(* IEC 61131-3 sources: mapprobotics-sample-tracking/FileDevices/GCode, 6 files *)

(* ---- ProdDetails.typ ---- *)
TYPE
	ProductDetailsType : 	STRUCT  (*Additional data added as attributes to every tracking object*)
		This : UDINT; (*Adress to the memory - debugging*)
		GripperClosed : BOOL; (*Gripper is close, product in manipulation*)
		TrackingFrameID : UDINT; (*tracking frame id*)
		PickPosDelta : McPosType;
		PickPos : McPosType; (*position where gripper has been closed*)
		IncrementPos : McPosType; (*change in position on frame*)
		Pos : McPosType; (*Actual Position of object*)
		ObjectType : USINT; (*Classification of the object (red / blue)*)
		InTracking : BOOL; (*Object is now active in Tracking*)
		Robot : DevicesListEnum; (*type of robot manipulated the object*)
	END_STRUCT;
	DevicesListEnum :
		( (*device definition of manipulating robots and axis*)
		DEV_Conveyor := 0, (*object id for conveyor*)
		DEV_Robot := 1, (*id for robot 1*)
		DEV_Removed := 2 (*marked as removed and do not show in scene*)
		);
END_TYPE

(* ---- Multipick.st ---- *)
#include 'ProdDetails.typ'

////////////////////////////////////////////////////////////////////////////////////
// INPUT Variables - configured as Program Elements of the interpreter
	// NextTrackingObjectIn : UDINT;							 Pointer to next object (GCS)

// OUTPUT Variables - configured as Program Elements of the interpreter
	// MaxPickPosIn : LREAL;								 	Maximum Position where robot is able to grab something (BCS)
	// MinPickPosIn : LREAL;								 	Minimum Position where objects are given to the robot (BCS)

VAR CONSTANT
	UpperZLevel : LREAL := 100.0;	// Gripper up position
	LowerZLevel : LREAL := 0.0;		// Gripper down position
	YProductPos : LREAL := 200;		// position in y coordinate where the product should be placed
END_VAR

VAR
	ActObj 	: REFERENCE TO ProductDetailsType;
	NextObj : REFERENCE TO ProductDetailsType;
	ParkPos				: McPointType := (Pos:=(X:=	  0, Y:= 0, 			Z:= UpperZLevel));
	SynchPosUp1			: McPointType := (Pos:=(X:=   -100, Y:= 0, 			Z:= UpperZLevel));
	SynchPosUp2			: McPointType := (Pos:=(X:=   100, Y:= 0, 			Z:= UpperZLevel));
	SynchPosDown1		: McPointType := (Pos:=(X:=   -100, Y:= 0, 			Z:= LowerZLevel));
	SynchPosDown2		: McPointType := (Pos:=(X:=   100, Y:= 0, 			Z:= LowerZLevel));
	StaticMoveDown		: McPointType := (Pos:=(X:=	  0, Y:= 0, 			Z:= 0));
	MoveToPark : BOOL 	:= FALSE;
END_VAR

PROGRAM _MAIN

	// Position init, reset frame in case of restart
	SetPCS(MachineFrame);
	MoveLR(ParkPos);

	// Set the manipulation area of the Robot
	MaxPickPosIn := 1400;
	MinPickPosIn := 200;

	REPEAT
		IF NextTrackingObjectIn <> 0 THEN
			MoveToPark := FALSE;

			ActObj ACCESS NextTrackingObjectIn;								// select the product
			TrackObjectR(ActObj.TrackingFrameID, SynchPosUp2, 50, 50);		// track on product
			MoveLR(SynchPosDown2);											// move to the take position
			SetM(34);														// Scene - remove product from belt, Close the gripper here
			WaitTime(0.04);													// Wait cause delay of gripper
			WaitALAP();
			MoveLR(SynchPosUp2);											// move up to change position

			NextObj ACCESS NextTrackingObjectIn;
			IF ADR(NextObj) <> 0 AND ADR(NextObj) <> ADR(ActObj) THEN
				TrackObjectR(NextObj.TrackingFrameID, SynchPosUp1, 50, 50);	// track on product
				MoveLR(SynchPosDown1);										// move to the take position
				SetM(33);													// Scene - remove product from belt, Close the gripper here
				WaitTime(0.04);												// Wait cause delay of gripper
				MoveLR(SynchPosUp1);										// move up to change position
			END_IF

			TrackStopR(FixedPlace, ParkPos, 50, 50);						// Move to the fixed place Position
			MoveLR(StaticMoveDown);											// move to the take position
			SetM(16);														// open the gripper here
			SetM(17);														// open the gripper here
			WaitTime(0.04);													// Wait cause delay of gripper
			MoveLR(ParkPos);												// move to the take position
			WaitALAP();

			IF NextTrackingObjectIn = 0 THEN								// Need to stop, no objects left
				MoveToPark := TRUE;											// force park position
			END_IF

		ELSE
			MoveToPark := TRUE;												// force park position, there is nothing to take
		END_IF

		IF MoveToPark THEN
			MoveLR(ParkPos);												// move to static park position
			WaitEndMove();													// sync interpreter and program
			WaitIp();														// hold interpreter until a new frame is available
		END_IF

	UNTIL FALSE END_REPEAT;

END_PROGRAM

(* ---- PickNPlace.st ---- *)
#include 'ProdDetails.typ'

////////////////////////////////////////////////////////////////////////////////////
// INPUT Variables - configured as Program Elements of the interpreter
	// NextTrackingObjectIn : UDINT;							 Pointer to next object (GCS)
	// NextTrackingObjectOut : UDINT;							 Pointer to next object (GCS)

// OUTPUT Variables - configured as Program Elements of the interpreter
	// MaxPickPosIn : LREAL;								 	Maximum Position where robot is able to grab something (BCS)
	// MinPickPosIn : LREAL;								 	Minimum Position where objects are given to the robot (BCS)
	// MaxPickPosOut : LREAL;								 	Maximum Position where robot is able to place something (BCS)
	// MinPickPosOut : LREAL;								 	Minimum Position where objects are placed by the robot (BCS)

VAR CONSTANT
	UpperZLevel : LREAL := 100.0;	// Gripper up position
	LowerZLevel : LREAL := 0.0;		// Gripper down position
	YProductPos : LREAL := 200;		// position in y coordinate where the product should be placed
END_VAR

VAR
	ActObj : REFERENCE TO ProductDetailsType;
	ParkPos				: McPointType := (Pos:=(X:=-100, Y:=100, 			Z:= UpperZLevel));
	SynchPosUp			: McPointType := (Pos:=(X:=   0, Y:= 0, 			Z:= UpperZLevel));
	SynchPosDown		: McPointType := (Pos:=(X:=   0, Y:= 0, 			Z:= LowerZLevel));
	MoveToPark : BOOL := FALSE;
END_VAR

PROGRAM _MAIN

	// Position init, reset frame in case of restart
	SetPCS(MachineFrame);
	MoveLR(ParkPos);

	// Set the manipulation area of the Robot
	MaxPickPosIn := 1400;
	MinPickPosIn := 400;
	MaxPickPosOut := 1700;
	MinPickPosOut := 700;

	REPEAT
		IF NextTrackingObjectIn <> 0 THEN
			MoveToPark := FALSE;

			ActObj ACCESS NextTrackingObjectIn;							// select the product
			TrackObjectR(ActObj.TrackingFrameID, SynchPosUp, 50, 50);	// track on product
			MoveLR(SynchPosDown);										// move to the take position
			WaitALAP();													// hold interpreter
			SetM(32);													// Scene - remove product from belt, close gripper
			WaitTime(0.04);												// Wait cause delay of gripper

			MoveLR(SynchPosUp);											// move up to change frame
			WaitUntil(NextTrackingObjectOut <> 0);						// hold interpeter until place frame has been selected
			ActObj ACCESS NextTrackingObjectOut;						// change memory reference
			TrackObjectR(ActObj.TrackingFrameID, SynchPosUp, 50, 50);	// move to place position
			MoveLR(SynchPosDown);										// move down on place position
			WaitALAP();													// hold interpreter
			SetM(16);													// Scene - place product on belt, open gripper
			WaitTime(0.04);												// Wait cause delay of gripper

			MoveLR(SynchPosUp);											// move up to change frame
			IF NextTrackingObjectIn = 0 THEN							// Need to stop, no objects left
				TrackStopR(MachineFrame, ParkPos, 50, 50);				// Move to a static frame
				MoveToPark := TRUE;										// force park position
			END_IF

		ELSE
			MoveToPark := TRUE;											// force park position, there is nothing to take
		END_IF

		IF MoveToPark THEN
			MoveLR(ParkPos);											// move to static park position
			WaitEndMove();												// sync interpreter and program
			WaitIp();													// hold interpreter until a new frame is available
		END_IF

	UNTIL FALSE END_REPEAT;

END_PROGRAM

(* ---- PlaceWithConditionalStop.st ---- *)
#include 'ProdDetails.typ'

////////////////////////////////////////////////////////////////////////////////////
// INPUT Variables - configured as Program Elements of the interpreter
	// NextTrackingObjectIn : UDINT;							 Pointer to next object (GCS)

// OUTPUT Variables - configured as Program Elements of the interpreter
	// MaxPickPosIn : LREAL;								 	Maximum Position where robot is able to grab something (BCS)
	// MinPickPosIn : LREAL;								 	Minimum Position where objects are given to the robot (BCS)

VAR CONSTANT
	UpperZLevel : LREAL := 100.0;	// Gripper up position
	LowerZLevel : LREAL := 0.0;		// Gripper down position
	YProductPos : LREAL := 200;		// position in y coordinate where the product should be placed
END_VAR

VAR
	ActObj : REFERENCE TO ProductDetailsType;
	ParkPos				: McPointType := (Pos:=(X:=	  0, Y:= 0, 			Z:= UpperZLevel));
	SynchPosUp			: McPointType := (Pos:=(X:=   0, Y:= 0, 			Z:= UpperZLevel));
	SynchPosDown		: McPointType := (Pos:=(X:=   0, Y:= 0, 			Z:= LowerZLevel));
	StaticMoveDown		: McPointType := (Pos:=(X:=   0, Y:= 0, 			Z:= -100));
	StaticMoveUp		: McPointType := (Pos:=(X:=   0, Y:= 0, 			Z:= 100));
	MoveToPark : BOOL 	:= FALSE;
END_VAR

PROGRAM _MAIN

	// Position init, reset frame in case of restart
	SetPCS(MachineFrame);
	MoveLR(ParkPos);

	// Set the manipulation area of the Robot
	MaxPickPosIn := 1400;
	MinPickPosIn := 200;

	REPEAT
		IF NextTrackingObjectIn <> 0 THEN
			MoveToPark := FALSE;

			ActObj ACCESS NextTrackingObjectIn;							// select the product
			TrackObjectR(ActObj.TrackingFrameID, SynchPosUp, 50, 50);	// track on product
			MoveLR(SynchPosDown);										// move to the take position
			// Close the gripper here
			SetM(32);													// Scene - remove product from belt
			WaitTime(0.04);												// Wait until gripper closes
			MoveLR(SynchPosUp);											// move up to change position

			TrackStopR(FixedPlace, ParkPos, 50, 50);					// Move to the fixed place Position
			ConditionalStop(123);										// Stop movement if place position is not valid
			Relative();													// use relative positions
			MoveLR(StaticMoveDown);										// move to the take position
			WaitEndMove();												// wait to go on with interpreter here
			SetM(16);													// open the gripper here
			WaitTime(0.04);												// Wait until gripper opens
			MoveLR(StaticMoveUp);										// move to the take position
			Absolute();

			IF NextTrackingObjectIn = 0 THEN							// Need to stop, no objects left
				MoveToPark := TRUE;										// force park position
			END_IF

		ELSE
			MoveToPark := TRUE;											// force park position, there is nothing to take
		END_IF

		IF MoveToPark THEN
			MoveLR(ParkPos);											// move to static park position
			WaitEndMove();												// sync interpreter and program
			WaitIp();													// hold interpreter until a new frame is available
		END_IF

	UNTIL FALSE END_REPEAT;

END_PROGRAM

(* ---- PrePalletizing.st ---- *)
#include 'ProdDetails.typ'

////////////////////////////////////////////////////////////////////////////////////
// INPUT Variables - configured as Program Elements of the interpreter
	// NextTrackingObjectIn : UDINT;							 Pointer to next object (GCS)

// OUTPUT Variables - configured as Program Elements of the interpreter
	// MaxPickPosIn : LREAL;								 	Maximum Position where robot is able to grab something (BCS)
	// MinPickPosIn : LREAL;								 	Minimum Position where objects are given to the robot (BCS)

VAR CONSTANT
	UpperZLevel : LREAL := 150.0;	// Gripper up position
	LowerZLevel : LREAL := 0.0;		// Gripper down position
	YProductPos : LREAL := 200;		// position in y coordinate where the product should be placed

	xStep : LREAL := 0.0;					// step size to get a tangential step for tracking
	yStep : LREAL := 0.1;					// step size to get a tangential step for tracking

END_VAR

VAR
	ActObj : REFERENCE TO ProductDetailsType;
	ParkPos						: McPointType := (Pos:=(X:=-350, 		Y:=-200, 			Z:= UpperZLevel));

	PreSynchPosUp				: McPointType := (Pos:=(X:=   0+xStep, 	Y:= 0+yStep, 		Z:= UpperZLevel));
	SynchPosUp					: McPointType := (Pos:=(X:=   0, 		Y:= 0, 				Z:= UpperZLevel));
	SynchPosDown				: McPointType := (Pos:=(X:=   0, 		Y:= 0, 				Z:= LowerZLevel));
	SynchPosForward				: McPointType := (Pos:=(X:= 100, 		Y:= 0, 				Z:= LowerZLevel));
	SynchPosSideward			: McPointType := (Pos:=(X:= 100, 		Y:= 100, 			Z:= LowerZLevel));
	SynchPosUpSideward			: McPointType := (Pos:=(X:= 100, 		Y:= 100, 			Z:= UpperZLevel));
	PostSynchPosUpSideward		: McPointType := (Pos:=(X:= 100-xStep, 	Y:=100-yStep,		Z:= UpperZLevel));

	MoveToPark : BOOL := FALSE;
	r1 : LREAL := 20.0;
END_VAR

// The radius is calculate by the half distance between two points this gives the result of a smooth interpolation
FUNCTION getRadius : LREAL
	VAR_INPUT
		posA : LREAL;
	END_VAR
	getRadius := MAX(20.0, ABS(posA) / 2.0);
END_FUNCTION

PROGRAM _MAIN

	EVAL('SERVICE_DATA["EXTENDED_TFA OFF"]', LANGUAGE_BR_GCODE);

	// Position init, reset frame in case of restart
	SetPCS(MachineFrame);
	MoveLR(ParkPos);

	// Set the manipulation area of the Robot
	MaxPickPosIn := 1400;
	MinPickPosIn := 1100;

	REPEAT
		IF NextTrackingObjectIn <> 0 THEN
			MoveToPark := FALSE;
			ActObj ACCESS NextTrackingObjectIn;							// select the product

			Feedrate(50000);
			r1 := getRadius(ActObj.Pos.Y);

			PreSynchPosUp := SynchPosUp;
			PostSynchPosUpSideward := SynchPosUpSideward;
			IF ActObj.Pos.Y > 0 THEN
				PreSynchPosUp.Pos.Y := PreSynchPosUp.Pos.Y - yStep;
				PostSynchPosUpSideward.Pos.Y := PostSynchPosUpSideward.Pos.Y - yStep;
			ELSE
				PreSynchPosUp.Pos.Y := PreSynchPosUp.Pos.Y + yStep;
				PostSynchPosUpSideward.Pos.Y := PostSynchPosUpSideward.Pos.Y + yStep;
			END_IF

			TrackObjectR(ActObj.TrackingFrameID, PreSynchPosUp, r1, r1);	// track on product
			MoveL(SynchPosUp);
			MoveLR(SynchPosDown);										// move to the take position

			SetM(8);													// Scene - start moving the poduct on the belt
			WaitTime(0.04);												// Wait cause delay of gripper
			Feedrate(15000);											// manipulate with reduced feedrate
			MoveL(SynchPosForward);										// move forward on belt
			MoveL(SynchPosSideward);									// move sideward on belt

			WaitALAP();													// hold interpreter
			// open the gripper here
			SetM(16);													// Scene - end of moving the product
			WaitTime(0.04);												// Wait cause delay of gripper
			MoveLR(SynchPosUpSideward);									// move up to change frame
			MoveLR(PostSynchPosUpSideward);									// move up to change frame

			IF NextTrackingObjectIn = 0 THEN							// Need to stop, no objects left
				TrackStopR(MachineFrame, ParkPos, 50, 50);				// Move to a static frame
				MoveToPark := TRUE;										// force park position
			END_IF

		ELSE
			MoveToPark := TRUE;											// force park position, there is nothing to take
		END_IF

		IF MoveToPark THEN
			MoveLR(ParkPos);											// move to static park position
			WaitEndMove();												// sync interpreter and program
			WaitIp();													// hold interpreter until a new frame is available
		END_IF

	UNTIL FALSE END_REPEAT;

END_PROGRAM

(* ---- Sorting.st ---- *)
#include 'ProdDetails.typ'

////////////////////////////////////////////////////////////////////////////////////
// INPUT Variables - configured as Program Elements of the interpreter
	// NextTrackingObjectIn : UDINT;							 Pointer to next object (GCS)
	// NextTrackingObjectOut : UDINT;							 Pointer to next object (GCS)

// OUTPUT Variables - configured as Program Elements of the interpreter
	// MaxPickPosIn : LREAL;								 	Maximum Position where robot is able to grab something (BCS)
	// MinPickPosIn : LREAL;								 	Minimum Position where objects are given to the robot (BCS)
	// MaxPickPosOut : LREAL;								 	Maximum Position where robot is able to place something (BCS)
	// MinPickPosOut : LREAL;								 	Minimum Position where objects are placed by the robot (BCS)

VAR CONSTANT
	UpperZLevel : LREAL := 100.0;	// Gripper up position
	LowerZLevel : LREAL := 0.0;		// Gripper down position
	YProductPos : LREAL := 200;		// position in y coordinate where the product should be placed
END_VAR

VAR
	ActObj : REFERENCE TO ProductDetailsType;
	ParkPos				: McPointType := (Pos:=(X:=	  0, Y:= 0, 			Z:= UpperZLevel));
	SynchPosUp			: McPointType := (Pos:=(X:=   0, Y:= 0, 			Z:= UpperZLevel));
	SynchPosDown		: McPointType := (Pos:=(X:=   0, Y:= 0, 			Z:= LowerZLevel));
	StaticMoveDown		: McPointType := (Pos:=(X:=	  0, Y:= 0, 			Z:= 0));
	MoveToPark : BOOL := FALSE;
END_VAR

PROGRAM _MAIN

	// Position init, reset frame in case of restart
	SetPCS(MachineFrame);
	MoveLR(ParkPos);

	// Set the manipulation area of the Robot
	MaxPickPosIn := 1400;
	MinPickPosIn := 400;
	MaxPickPosOut := 1700;
	MinPickPosOut := 700;

	REPEAT
		IF NextTrackingObjectIn <> 0 THEN
			MoveToPark := FALSE;

			ActObj ACCESS NextTrackingObjectIn;								// select the product
			TrackObjectR(ActObj.TrackingFrameID, SynchPosUp, 50, 50);		// track on product
			MoveLR(SynchPosDown);											// move to the take position
			WaitALAP();														// hold interpreter
			// Close the gripper here
			SetM(32);														// Scene - remove product from belt
			WaitTime(0.04);													// Wait until gripper opens
			MoveLR(SynchPosUp);												// move up to change frame

			IF ActObj.ObjectType = 1 THEN									// sort out objects of type 1
				TrackStopR(FixedPlace, ParkPos, 50, 50);					// Move to the fixed place Position
				MoveLR(StaticMoveDown);										// move to the take position
				SetM(16);													// open the gripper here
				WaitTime(0.04);												// Wait until gripper opens
				MoveLR(ParkPos);											// move to the take position
				WaitALAP();

				IF NextTrackingObjectIn = 0 THEN							// Need to stop, no objects left
					MoveToPark := TRUE;										// force park position
				END_IF

			ELSE

				WaitUntil(NextTrackingObjectOut <> 0);						// hold interpeter until place frame has been selected
				ActObj ACCESS NextTrackingObjectOut;						// change memory reference
				TrackObjectR(ActObj.TrackingFrameID, SynchPosUp, 50, 50);	// move to place position
				MoveLR(SynchPosDown);										// move down on place position
				WaitALAP();													// hold interpreter
				ActObj.ObjectType := 0;										// set type of object (scene generation)
				SetM(16);													// Scene - place product on belt, Open the gripper here
				WaitTime(0.04);												// Wait until gripper opens
				MoveLR(SynchPosUp);											// move up to change frame
				IF NextTrackingObjectIn = 0 THEN							// Need to stop, no objects left
					TrackStopR(MachineFrame, ParkPos, 50, 50);				// Move to a static frame
					MoveToPark := TRUE;										// force park position
				END_IF
			END_IF

		ELSE
			MoveToPark := TRUE;											// force park position, there is nothing to take
		END_IF

		IF MoveToPark THEN
			MoveLR(ParkPos);											// move to static park position
			WaitEndMove();												// sync interpreter and program
			WaitIp();													// hold interpreter until a new frame is available
		END_IF

	UNTIL FALSE END_REPEAT;

END_PROGRAM
